// TIA Portal V20 export
TYPE "Kistler_Dateinamen_ges"
   STRUCT
      Kistler_Dateinamen_ges : Array[0..59] of Char;
   END_STRUCT;
END_TYPE
